{attribute 'pack_mode' := '1'}
TYPE ST_EssPublish_V1 :
STRUCT
	DeviceIndex	:	UDINT;
	Status	:	UDINT;
	AcActivePower	:	REAL;
	AcReactivePower:	REAL;
	AcVoltageR     :	REAL;
	AcVoltageS     :	REAL;
	AcVoltageT     :	REAL;
	AcCurrentR     :	REAL;
	AcCurrentS     :	REAL;
	AcCurrentT     :	REAL;
	Frequency      :	REAL;
	PowerFactor    :	REAL;
	EnergyActivePower:	REAL;
	EnergyReactivePower:	REAL;
	EnergyReverseActivePower:	REAL;
	EnergyReverseReactivePower:	REAL;
	Warning1:	UDINT;
	Warning2:	UDINT;
	Warning3:	UDINT;
	Warning4:	UDINT;
	Warning5:	UDINT;
	Warning6:	UDINT;
	Warning7:	UDINT;
	Warning8:	UDINT;
	Warning9:	UDINT;
	Warning10:	UDINT;
	Fault1:		UDINT;
	Fault2:		UDINT;
	Fault3:		UDINT;
	Fault4:		UDINT;
	Fault5:		UDINT;
	Fault6:		UDINT;
	Fault7:		UDINT;
	Fault8:		UDINT;
	Fault9:		UDINT;
	Fault10:		UDINT;
END_STRUCT
END_TYPE

(* stored: Version 1.1.0.1, ProductVersion 3.1.4024.9
   DUT ST_EssPublish_V1: Id {6662cbf1-6ddf-4e3e-9d52-ec7ae570071a} *)
